(* IEC 61131-3 sources: platen-temp-control/plc, 4 files *)

(* ---- FB_PI_AntiWindup.st ---- *)
(* FB_PI_AntiWindup
   Discrete PI controller with clamping anti-windup and bumpless manual mode.
   Same algorithm as matlab/sim_pi.m, so simulation and PLC results match.
   Call once every Ts seconds (e.g., every 10th scan of a 100 ms task). *)
FUNCTION_BLOCK FB_PI_AntiWindup
VAR_INPUT
    xEnable    : BOOL;            (* TRUE = control, FALSE = output 0 and reset *)
    xManual    : BOOL;            (* TRUE = manual mode *)
    rManualOut : REAL;            (* manual output 0..1 *)
    rSP        : REAL;            (* setpoint [degC] *)
    rPV        : REAL;            (* process value [degC] *)
    rKp        : REAL := 0.0486;  (* proportional gain [1/degC] *)
    rTi        : REAL := 288.0;   (* integral time [s] *)
    rTs        : REAL := 1.0;     (* sample time [s] *)
    rOutMin    : REAL := 0.0;
    rOutMax    : REAL := 1.0;
    xAntiWindup: BOOL := TRUE;    (* set FALSE to demonstrate windup *)
END_VAR
VAR_OUTPUT
    rOut       : REAL;            (* controller output 0..1 *)
    rError     : REAL;
    xSaturated : BOOL;
END_VAR
VAR
    rI         : REAL;            (* integral term *)
    rOutRaw    : REAL;
    xPushHigh  : BOOL;
    xPushLow   : BOOL;
END_VAR

IF NOT xEnable THEN
    rI := 0.0;
    rOut := 0.0;
    xSaturated := FALSE;
    RETURN;
END_IF

rError := rSP - rPV;

IF xManual THEN
    rOut := LIMIT(rOutMin, rManualOut, rOutMax);
    (* bumpless transfer: preload integral so auto starts from manual output *)
    rI := rOut - rKp * rError;
    RETURN;
END_IF

rOutRaw := rKp * rError + rI;
rOut := LIMIT(rOutMin, rOutRaw, rOutMax);

xPushHigh := (rOutRaw > rOutMax) AND (rError > 0.0);
xPushLow  := (rOutRaw < rOutMin) AND (rError < 0.0);
xSaturated := xPushHigh OR xPushLow;

IF (NOT xAntiWindup) OR (NOT xSaturated) THEN
    IF rTi > 0.0 THEN
        rI := rI + rKp * rTs / rTi * rError;
    END_IF
END_IF
END_FUNCTION_BLOCK

(* ---- FB_PlatenModel.st ---- *)
(* FB_PlatenModel
   Simulated heater + platen (same equations as matlab/platen_params.m).
   Lets the soft PLC run a full test with no hardware.
   Forward Euler integration; keep rDt <= 0.5 s (fast heater time constant ~8 s). *)
FUNCTION_BLOCK FB_PlatenModel
VAR_INPUT
    rU      : REAL;            (* heater command 0..1 *)
    rW      : REAL;            (* disturbance heat [W], negative = cold mold *)
    rDt     : REAL := 0.1;     (* integration step = task cycle [s] *)
    xReset  : BOOL;            (* TRUE = back to ambient *)
END_VAR
VAR_OUTPUT
    rTh     : REAL := 25.0;    (* heater temperature [degC] *)
    rTp     : REAL := 25.0;    (* platen temperature [degC] *)
END_VAR
VAR
    rCh     : REAL := 800.0;
    rCp     : REAL := 14000.0;
    rRhp    : REAL := 0.01;
    rRpa    : REAL := 0.155;
    rPmax   : REAL := 4000.0;
    rTa     : REAL := 25.0;
    rQhp    : REAL;            (* heat flow heater -> platen [W] *)
    rQloss  : REAL;            (* heat loss platen -> ambient [W] *)
END_VAR

IF xReset THEN
    rTh := rTa;
    rTp := rTa;
    RETURN;
END_IF

rQhp   := (rTh - rTp) / rRhp;
rQloss := (rTp - rTa) / rRpa;
rTh := rTh + rDt * (rPmax * LIMIT(0.0, rU, 1.0) - rQhp) / rCh;
rTp := rTp + rDt * (rQhp - rQloss + rW) / rCp;
END_FUNCTION_BLOCK

(* ---- FB_TimeProportional.st ---- *)
(* FB_TimeProportional
   Turns a 0..1 duty into an ON/OFF output for a solid-state relay (SSR).
   Example: rDuty = 0.3, cycle 2 s -> ON 0.6 s, OFF 1.4 s. *)
FUNCTION_BLOCK FB_TimeProportional
VAR_INPUT
    rDuty   : REAL;            (* 0..1 *)
    tCycle  : TIME := T#2S;    (* SSR cycle time *)
END_VAR
VAR_OUTPUT
    xOut    : BOOL;            (* wire to the SSR output card *)
END_VAR
VAR
    fbCycle : TON;
    tOn     : TIME;
END_VAR

fbCycle(IN := NOT fbCycle.Q, PT := tCycle);
tOn := REAL_TO_TIME(LIMIT(0.0, rDuty, 1.0) * TIME_TO_REAL(tCycle));
xOut := fbCycle.ET < tOn;
END_FUNCTION_BLOCK

(* ---- PLC_PRG.st ---- *)
(* PLC_PRG  -  run in a cyclic task at 100 ms.
   Heat-up, PI control every 1 s, over-temperature and sensor-fault trips,
   and a cold-mold disturbance button for testing. Values in degC (177 C = 350 F). *)
PROGRAM PLC_PRG
VAR
    (* operator / HMI *)
    xStart          : BOOL;
    xStop           : BOOL;
    xResetAlarm     : BOOL;
    xLoadColdMold   : BOOL;            (* HMI test button *)
    xManual         : BOOL;
    rManualOut      : REAL;
    rSetpoint       : REAL := 177.0;
    rHighLimit      : REAL := 190.0;   (* over-temperature trip *)

    (* state *)
    xRunning        : BOOL;
    xAlarmOverTemp  : BOOL;
    xAlarmSensor    : BOOL;
    xAtTemp         : BOOL;            (* within +/-2 C: ready to cure *)

    (* simulation *)
    xSimulate       : BOOL := TRUE;    (* FALSE = use the real sensor input *)
    rRealPV         : REAL;            (* map to the analog input card *)
    rPV             : REAL;
    rDisturbanceW   : REAL;
    fbMold          : TP;

    (* blocks *)
    fbPI            : FB_PI_AntiWindup;
    fbPlant         : FB_PlatenModel;
    fbSSR           : FB_TimeProportional;
    xHeaterOut      : BOOL;            (* map to the SSR digital output *)
    iScan           : INT;
    rDuty           : REAL;
    fbAtTemp        : TON;
END_VAR

(* ---- start / stop ---- *)
IF xStop OR xAlarmOverTemp OR xAlarmSensor THEN
    xRunning := FALSE;
ELSIF xStart THEN
    xRunning := TRUE;
END_IF

(* ---- measurement ---- *)
IF xSimulate THEN
    rPV := fbPlant.rTp;
ELSE
    rPV := rRealPV;
END_IF

(* ---- trips (latched until reset) ---- *)
IF rPV > rHighLimit THEN xAlarmOverTemp := TRUE; END_IF
IF (rPV < -20.0) OR (rPV > 400.0) THEN xAlarmSensor := TRUE; END_IF
IF xResetAlarm AND (rPV < rHighLimit - 5.0) AND (rPV > -20.0) AND (rPV < 400.0) THEN
    xAlarmOverTemp := FALSE;
    xAlarmSensor := FALSE;
END_IF

(* ---- PI controller every 10 scans = 1 s ---- *)
iScan := iScan + 1;
IF iScan >= 10 THEN
    iScan := 0;
    fbPI(xEnable := xRunning, xManual := xManual, rManualOut := rManualOut,
         rSP := rSetpoint, rPV := rPV, rTs := 1.0);
    rDuty := fbPI.rOut;
END_IF
IF NOT xRunning THEN rDuty := 0.0; END_IF

(* ---- heater output ---- *)
fbSSR(rDuty := rDuty, tCycle := T#2S);
xHeaterOut := fbSSR.xOut AND xRunning;

(* ---- at-temperature indication (stable 30 s) ---- *)
fbAtTemp(IN := xRunning AND (ABS(rSetpoint - rPV) <= 2.0), PT := T#30S);
xAtTemp := fbAtTemp.Q;

(* ---- simulated plant + cold-mold disturbance (90 s, -3000 W) ---- *)
fbMold(IN := xLoadColdMold, PT := T#90S);
IF fbMold.Q THEN rDisturbanceW := -3000.0; ELSE rDisturbanceW := 0.0; END_IF
(* the plant sees the averaged duty; use BOOL_TO_REAL(xHeaterOut) to see SSR ripple *)
fbPlant(rU := rDuty, rW := rDisturbanceW, rDt := 0.1);
END_PROGRAM
